Staubli VAL3: Init_Repere.pgx

program Init_Repere()
begin
  bInit_repere =true
  setFrame(pRcaisse[0], pRcaisse[1], pRcaisse[2],fcaisse)
end
